// TIA Portal V20 export
TYPE "MC_Variablen"
   STRUCT
      Antrieb_Ein : Struct
         Enable : Bool;
         StartMode : DInt;
         StopMode : Int;
         Status : Bool;
         Busy : Bool;
         Error : Bool;
         ErrorID : Word;
      END_STRUCT;
      Antieb_Reset : Struct
         Execute : Bool;
         Restart : Bool;
         Done : Bool;
         Busy : Bool;
         ComandAborted : Bool;
         Error : Bool;
         ErrorID : Word;
      END_STRUCT;
      Antrieb_Referenz : Struct
         Execute : Bool;
         Position : LReal;
         Mode : Int;
         ReferenceMarkPosition : LReal;
         Done : Bool;
         Busy : Bool;
         ComandAborted : Bool;
         Error : Bool;
         ErrorID : Word;
      END_STRUCT;
      Antrieb_Move_Absolute : Struct
         Execute : Bool;
         Position : LReal;
         Velocity : LReal;
         Acceleration : LReal;
         Deceleration : LReal;
         Jerk : LReal;
         Direction : Int;
         Done : Bool;
         Busy : Bool;
         ComandAborted : Bool;
         Error : Bool;
         ErrorID : Word;
      END_STRUCT;
   END_STRUCT;
END_TYPE
